// TIA Portal V20 export
DATA_BLOCK "HW_Status_DB"   // DB166
{ S7_Optimized_Access := 'TRUE' }
// stored: MemoryReserve 100
   VAR
      State : Array[0..1023] of Bool;
   END_VAR
BEGIN
   State[0..1023] := FALSE;
END_DATA_BLOCK
